(*
SPDX-License-Identifier: MIT
License: https://opensource.org/license/mit
*)

(*!
<summary>Owns an arithmetic test and a nested timing group.</summary>
<description>
Owns persistent child storage and fixed parent associations. Use in one task without reentry.
Children is borrowed and must not be modified by application code. Constructor callbacks are not used.
</description>
*)

{attribute 'no_assign'}
{attribute 'no_explicit_call' := 'do not call this function block directly'}
FUNCTION_BLOCK BasicTestGroup EXTENDS TOF_Testing.TestGroup<2>
VAR_STAT
	{attribute 'hide'}
	_ClassName : STRING := __POUNAME();
END_VAR
VAR
	_Addition : AdditionTest(name := "Addition", parent := THIS^);
	_Timing : TimingTestGroup(name := "Timing", parent := THIS^);

	_Children : ARRAY [0.._ChildCount - 1] OF TOF_Testing.ITestElement :=
	[
		_Addition,
		_Timing
	];
END_VAR

//! <summary>Borrows the fixed array of this concrete group; do not modify it.</summary>
{attribute 'monitoring' := 'call'}
PROPERTY Children : REFERENCE TO ARRAY [0.._ChildCount - 1] OF TOF_Testing.ITestElement
GET
Children REF= _Children;
END_GET
END_PROPERTY

//! <summary>Borrows the concrete class name for the lifetime of this instance; callers must not modify it.</summary>
{attribute 'monitoring' := 'call'}
PROPERTY ClassName : REFERENCE TO STRING
GET
ClassName REF= _ClassName;
END_GET
END_PROPERTY

//! <summary>Borrows the compiler-initialized namespace; callers must not modify the returned reference.</summary>
{attribute 'monitoring' := 'call'}
PROPERTY NamespaceName : REFERENCE TO STRING
GET
NamespaceName REF= CurrentNamespace.Name;
END_GET
END_PROPERTY

//! <summary>Reports the complete concrete instance size, excluding separately allocated storage.</summary>
{attribute 'monitoring' := 'call'}
PROPERTY SelfSize : ULINT
GET
SelfSize := XSIZEOF(THIS^);
END_GET
END_PROPERTY

END_FUNCTION_BLOCK

(* stored: Version 1.1.0.1
   POU BasicTestGroup: Id {42c98e9a-fb60-4225-918f-3a742a324332}, SpecialFunc None
   Property Children: Id {1ca423b8-e742-44d4-8d9f-eb2138ab07f1}
   Get Get: Id {cd89a098-d960-440c-98f7-0c79bb0bc818}
   Property ClassName: Id {23b902d9-a159-4a3d-960f-5ca4bfe5f1b9}
   Get Get: Id {672e4920-1fb2-4094-b742-6d7cfd8de785}
   Property NamespaceName: Id {09e25467-2cf2-4c61-b927-5f954614590a}
   Get Get: Id {421501c9-1501-4a9f-adf5-f0407d5aa687}
   Property SelfSize: Id {a5895aa0-5ff0-4a40-b2b4-7cbe25acf0c6}
   Get Get: Id {98cfb46b-c46d-42bf-9f5a-31ab7c7b4dc2} *)
